TYPE ST_PolarIIChamber_CleanSetting :
STRUCT
	TargetCupIndex : UINT; // 1..4
	CleanType : E_PolarIIChamberCleanType;
END_STRUCT
END_TYPE

(* stored: Version 1.1.0.1, ProductVersion 3.1.4026.18
   DUT ST_PolarIIChamber_CleanSetting: Id {14000000-0000-0000-0000-000000000009} *)
